FUNCTION_BLOCK FB_Register
VAR_INPUT
END_VAR
VAR_OUTPUT
END_VAR
VAR
	arrRegister     : ARRAY[1..100] OF ITF_Base;
    nNoOfInterfaces : UDINT := 0;
END_VAR

METHOD PUBLIC AddInterfacePointer : UDINT
VAR_INPUT
	ipBase : ITF_Base;
END_VAR
VAR
	n : UDINT;
END_VAR
// 0 bedeutet: Registrierung nicht erfolgreich.
AddInterfacePointer := 0;

// Eine leere Interface-Referenz nicht aufnehmen.
IF ipBase = 0 THEN
    RETURN;
END_IF

// Bereits registriert? Bestehenden Platz zurückgeben.
FOR n := 1 TO nNoOfInterfaces DO
    IF arrRegister[n] = ipBase THEN
        AddInterfacePointer := n;
        RETURN;
    END_IF
END_FOR

// Bei vollem Register nichts verändern.
IF nNoOfInterfaces >= 100 THEN
    RETURN;
END_IF

// Neue Referenz speichern.
nNoOfInterfaces := nNoOfInterfaces + 1;
arrRegister[nNoOfInterfaces] := ipBase;

// Zugewiesenen Tabellenplatz zurückgeben.
AddInterfacePointer := nNoOfInterfaces;
END_METHOD

END_FUNCTION_BLOCK

(* stored: Version 1.1.0.1, ProductVersion 3.1.4024.16
   POU FB_Register: Id {1592dd4e-b7ea-4f87-a486-63caf88324df}, SpecialFunc None
   Method AddInterfacePointer: Id {a647cf0f-ce03-4af8-a2f2-1948af184ec9} *)
